// TIA Portal V20 export
FUNCTION_BLOCK "PR_Gantry_2_Soft2.0 1_workflow_0f74f7"   // FB44, LAD
{ S7_Optimized_Access := 'TRUE' }
// stored: MemoryReserve 100, SetENOAutomatically false
   VAR_INPUT
      iAcceptPartPick : Bool;
      iAcceptPartPlace : Bool;
      iAutoRunning : Bool;
      iFaultReset : Bool;
      iFibroSafe : Bool;
      iOTS_Frm_Shuttle : Bool;
      iPartPresent : Bool;
      iPartPresent_Fibro : Bool;
      iPartUngrip : Bool;
      iRTR_Frm_Fibro : Bool;
      iReset_fault : Bool;
      iShuttleAtPickPos : Bool;
      iShuttleSafe : Bool;
      iSstMode : Bool;
      iSstPB : Bool;
      iXAxisAtPartPickPos : Bool;
      iXAxisAtPlacePos : Bool;
      iXAxisSafe : Bool;
      iZAxisDownPlace : Bool;
      iZAxisPickPos : Bool;
      iZAxisSafe : Bool;
      iZAxisUp : Bool;
   END_VAR
   VAR_OUTPUT
      qError : Array[0..8] of Bool;
      qMessage : Array[0..1] of Bool;
      qOTS_To_Fibro : Bool;
      qPartUngripCmd : Bool;
      qRTR_To_Shuttle : Bool;
      qXAxisHomeCmd : Bool;
      qXAxisHomeCmdPlace : Bool;
      qXAxisPickPosCmd : Bool;
      qZAxisDownCmd : Bool;
      qZAxisHomeCmd : Bool;
      qZAxisUpCmd : Bool;
      qZDownCmd : Bool;
   END_VAR
   VAR
      c170_ChkPartPlaced_T1 : Bool;
      c170_ChkPartPlaced_T2 : Bool;
      c180_WtOperatorDecisionPlace_T1 : Bool;
      c180_WtOperatorDecisionPlace_T2 : Bool;
      c40_ChkPartPresent_T1 : Bool;
      c40_ChkPartPresent_T2 : Bool;
      c40_ChkPartPresent_T3 : Bool;
      c90_ChkPartPick_T1 : Bool;
      c90_ChkPartPick_T2 : Bool;
      StateNo : Int;
      s100_WtOperatorDecision : Bool;
      s100_WtOperatorDecision_T1 : Bool;
      s100_WtOperatorDecision_T2 : Bool;
      s10_WtAllAtSafe : Bool;
      s10_WtAllAtSafe_T1 : Bool;
      s110_WtZAxisUp : Bool;
      s110_WtZAxisUp_T1 : Bool;
      s120_ChkFibroSafe : Bool;
      s120_ChkFibroSafe_T1 : Bool;
      s130_WtXAxisPlacePos : Bool;
      s130_WtXAxisPlacePos_T1 : Bool;
      s140_WtRTRFrmFibro : Bool;
      s140_WtRTRFrmFibro_T1 : Bool;
      s150_WtZAxisDownPlace : Bool;
      s150_WtZAxisDownPlace_T1 : Bool;
      s160_WtPartUngrip : Bool;
      s160_WtPartUngrip_T1 : Bool;
      s170_ChkPartPlaced : Bool;
      s170_ChkPartPlaced_T1 : Bool;
      s170_ChkPartPlaced_T2 : Bool;
      s180_WtOperatorDecisionPlace : Bool;
      s180_WtOperatorDecisionPlace_T1 : Bool;
      s180_WtOperatorDecisionPlace_T2 : Bool;
      s1_ResetRelease : Bool;
      s1_ResetRelease_T1 : Bool;
      s20_WtZAxisSafe : Bool;
      s20_WtZAxisSafe_T1 : Bool;
      s30_WtXAxisAtSafe : Bool;
      s30_WtXAxisAtSafe_T1 : Bool;
      s40_ChkPartPresent : Bool;
      s40_ChkPartPresent_T1 : Bool;
      s40_ChkPartPresent_T2 : Bool;
      s40_ChkPartPresent_T3 : Bool;
      s45_WtOperatorAck : Bool;
      s45_WtOperatorAck_T1 : Bool;
      s50_WtShuttleAtSafe : Bool;
      s50_WtShuttleAtSafe_T1 : Bool;
      s60_WtXAxisPickPos : Bool;
      s60_WtXAxisPickPos_T1 : Bool;
      s70_WtOTSFrmShuttle : Bool;
      s70_WtOTSFrmShuttle_T1 : Bool;
      s80_WtZAxisPickPos : Bool;
      s80_WtZAxisPickPos_T1 : Bool;
      s90_ChkPartPick : Bool;
      s90_ChkPartPick_T1 : Bool;
      s90_ChkPartPick_T2 : Bool;
      sAbnormalStatus : Bool;
      sPartPresentInGrip : Bool;
      sSst : Bool;
      sSstPulse : Bool;
      sSstRise : Bool;
      sStWtResetRel : Bool;
      sStWtResetRel_T1 : Bool;
   END_VAR
   VAR_TEMP
      tOne : Bool;
   END_VAR
   VAR_TEMP   // added for the SCL form of the ladder/FBD networks
      _w1 : Bool;
      _w2 : Bool;
   END_VAR
BEGIN

REGION Network 1
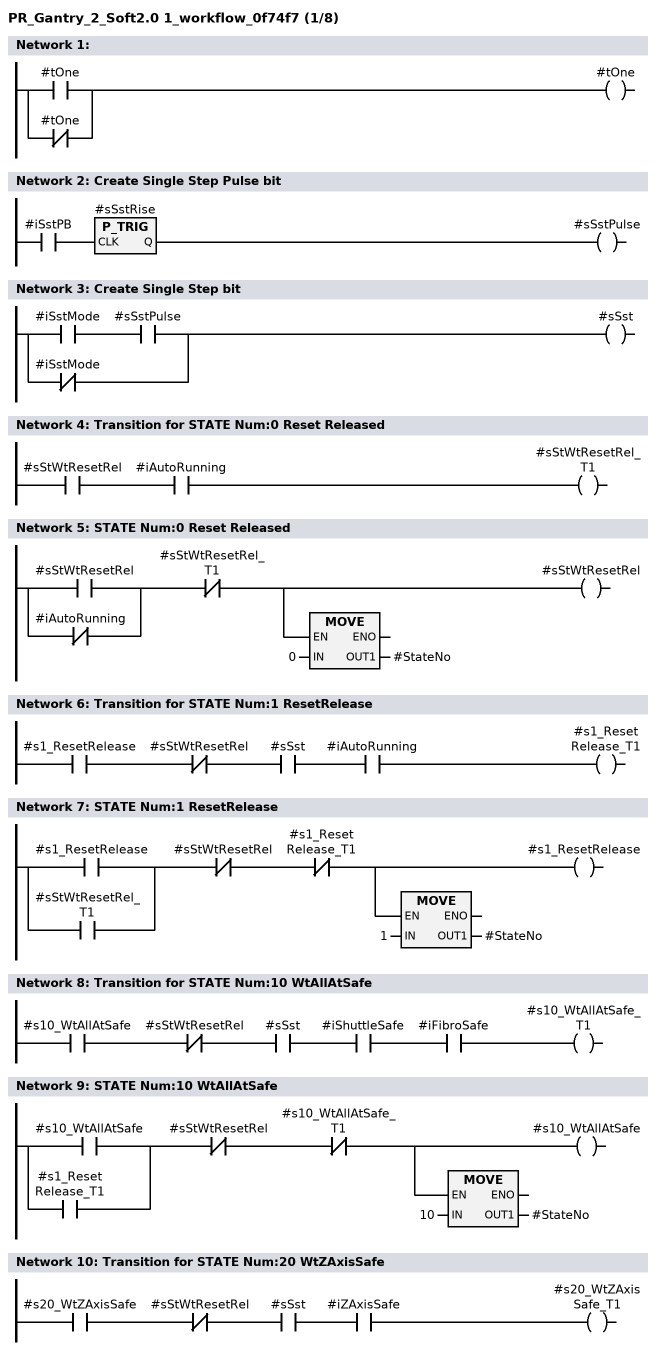
   RUNG wire#powerrail
      Contact( #tOne )
      wire#w1
      Coil( #tOne )
   END_RUNG
   RUNG wire#powerrail
      I_Contact( #tOne )
   END_RUNG wire#w1
   // the same network as SCL:
   #tOne := #tOne OR NOT #tOne;
END_REGION

REGION Network 2: Create Single Step Pulse bit
   RUNG wire#powerrail
      Contact( #iSstPB )
      P_Trig( #sSstRise )
      Coil( #sSstPulse )
   END_RUNG
   // the same network as SCL:
   #_w1 := #iSstPB AND NOT #sSstRise;   // rising edge
   #sSstRise := #iSstPB;
   #sSstPulse := #_w1;
END_REGION

REGION Network 3: Create Single Step bit
   RUNG wire#powerrail
      Contact( #iSstMode )
      Contact( #sSstPulse )
      wire#w1
      Coil( #sSst )
   END_RUNG
   RUNG wire#powerrail
      I_Contact( #iSstMode )
   END_RUNG wire#w1
   // the same network as SCL:
   #sSst := (#iSstMode AND #sSstPulse) OR NOT #iSstMode;
END_REGION

REGION Network 4: Transition for STATE Num:0 Reset Released
   RUNG wire#powerrail
      Contact( #sStWtResetRel )
      Contact( #iAutoRunning )
      Coil( #sStWtResetRel_T1 )
   END_RUNG
   // the same network as SCL:
   #sStWtResetRel_T1 := #sStWtResetRel AND #iAutoRunning;
END_REGION

REGION Network 5: STATE Num:0 Reset Released
   RUNG wire#powerrail
      Contact( #sStWtResetRel )
      wire#w1
      I_Contact( #sStWtResetRel_T1 )
      wire#w2
      Coil( #sStWtResetRel )
   END_RUNG
   RUNG wire#powerrail
      I_Contact( #iAutoRunning )
   END_RUNG wire#w1
   RUNG wire#w2
      { S7_GenerateENO := "TRUE" } Move(in := 0, out1 => #StateNo)
   END_RUNG
   // the same network as SCL:
   #sStWtResetRel := (#sStWtResetRel OR NOT #iAutoRunning) AND NOT #sStWtResetRel_T1;
   IF #sStWtResetRel THEN #StateNo := 0; END_IF;
END_REGION

REGION Network 6: Transition for STATE Num:1 ResetRelease
   RUNG wire#powerrail
      Contact( #s1_ResetRelease )
      I_Contact( #sStWtResetRel )
      Contact( #sSst )
      Contact( #iAutoRunning )
      Coil( #s1_ResetRelease_T1 )
   END_RUNG
   // the same network as SCL:
   #s1_ResetRelease_T1 := #s1_ResetRelease AND NOT #sStWtResetRel AND #sSst AND #iAutoRunning;
END_REGION

REGION Network 7: STATE Num:1 ResetRelease
   RUNG wire#powerrail
      Contact( #s1_ResetRelease )
      wire#w1
      I_Contact( #sStWtResetRel )
      I_Contact( #s1_ResetRelease_T1 )
      wire#w2
      Coil( #s1_ResetRelease )
   END_RUNG
   RUNG wire#powerrail
      Contact( #sStWtResetRel_T1 )
   END_RUNG wire#w1
   RUNG wire#w2
      { S7_GenerateENO := "TRUE" } Move(in := 1, out1 => #StateNo)
   END_RUNG
   // the same network as SCL:
   #s1_ResetRelease := (#s1_ResetRelease OR #sStWtResetRel_T1) AND NOT #sStWtResetRel AND NOT #s1_ResetRelease_T1;
   IF #s1_ResetRelease THEN #StateNo := 1; END_IF;
END_REGION

REGION Network 8: Transition for STATE Num:10 WtAllAtSafe
   RUNG wire#powerrail
      Contact( #s10_WtAllAtSafe )
      I_Contact( #sStWtResetRel )
      Contact( #sSst )
      Contact( #iShuttleSafe )
      Contact( #iFibroSafe )
      Coil( #s10_WtAllAtSafe_T1 )
   END_RUNG
   // the same network as SCL:
   #s10_WtAllAtSafe_T1 := #s10_WtAllAtSafe AND NOT #sStWtResetRel AND #sSst AND #iShuttleSafe AND #iFibroSafe;
END_REGION

REGION Network 9: STATE Num:10 WtAllAtSafe
   RUNG wire#powerrail
      Contact( #s10_WtAllAtSafe )
      wire#w1
      I_Contact( #sStWtResetRel )
      I_Contact( #s10_WtAllAtSafe_T1 )
      wire#w2
      Coil( #s10_WtAllAtSafe )
   END_RUNG
   RUNG wire#powerrail
      Contact( #s1_ResetRelease_T1 )
   END_RUNG wire#w1
   RUNG wire#w2
      { S7_GenerateENO := "TRUE" } Move(in := 10, out1 => #StateNo)
   END_RUNG
   // the same network as SCL:
   #s10_WtAllAtSafe := (#s10_WtAllAtSafe OR #s1_ResetRelease_T1) AND NOT #sStWtResetRel AND NOT #s10_WtAllAtSafe_T1;
   IF #s10_WtAllAtSafe THEN #StateNo := 10; END_IF;
END_REGION

REGION Network 10: Transition for STATE Num:20 WtZAxisSafe
   RUNG wire#powerrail
      Contact( #s20_WtZAxisSafe )
      I_Contact( #sStWtResetRel )
      Contact( #sSst )
      Contact( #iZAxisSafe )
      Coil( #s20_WtZAxisSafe_T1 )
   END_RUNG
   // the same network as SCL:
   #s20_WtZAxisSafe_T1 := #s20_WtZAxisSafe AND NOT #sStWtResetRel AND #sSst AND #iZAxisSafe;
END_REGION

REGION Network 11: STATE Num:20 WtZAxisSafe
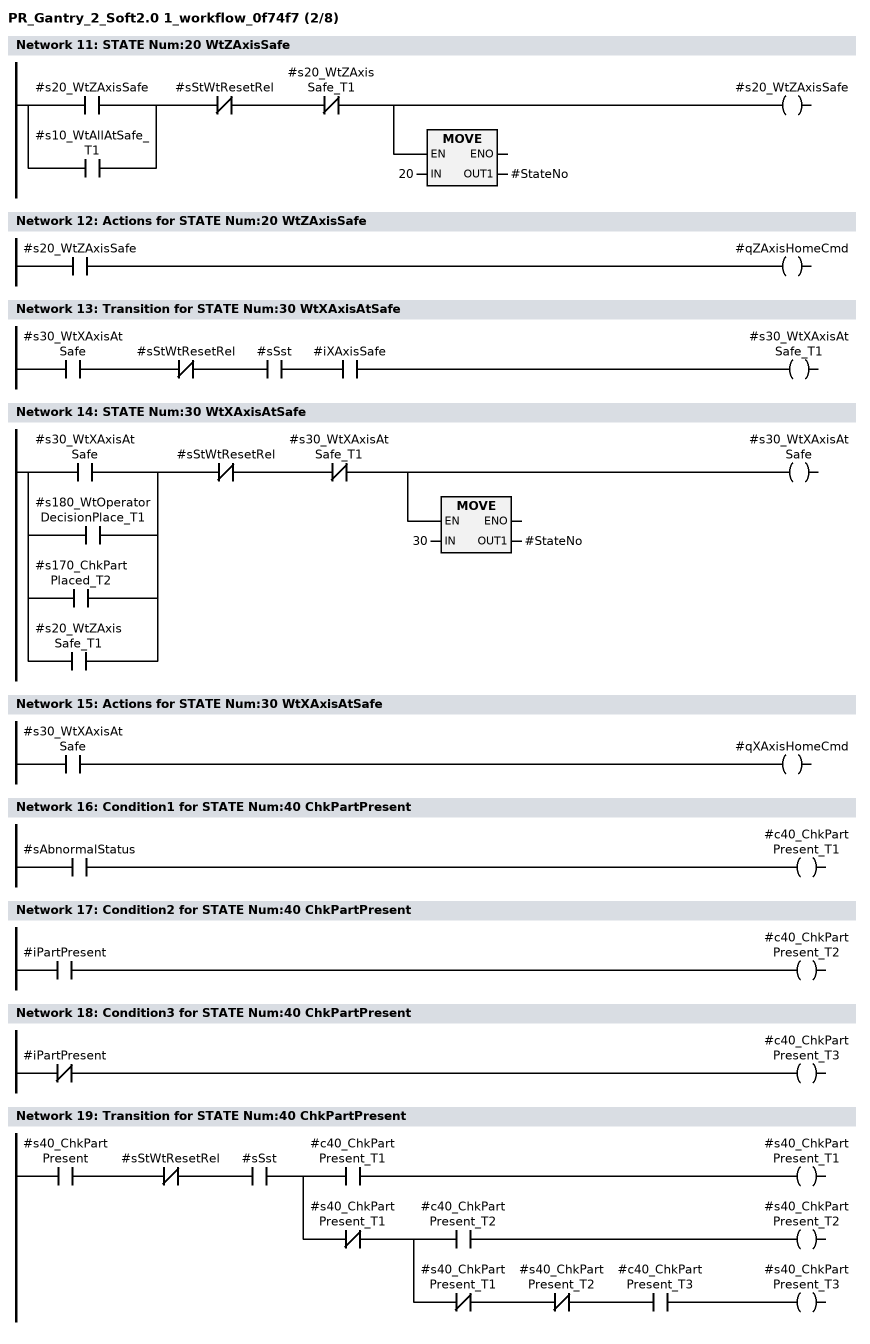
   RUNG wire#powerrail
      Contact( #s20_WtZAxisSafe )
      wire#w1
      I_Contact( #sStWtResetRel )
      I_Contact( #s20_WtZAxisSafe_T1 )
      wire#w2
      Coil( #s20_WtZAxisSafe )
   END_RUNG
   RUNG wire#powerrail
      Contact( #s10_WtAllAtSafe_T1 )
   END_RUNG wire#w1
   RUNG wire#w2
      { S7_GenerateENO := "TRUE" } Move(in := 20, out1 => #StateNo)
   END_RUNG
   // the same network as SCL:
   #s20_WtZAxisSafe := (#s20_WtZAxisSafe OR #s10_WtAllAtSafe_T1) AND NOT #sStWtResetRel AND NOT #s20_WtZAxisSafe_T1;
   IF #s20_WtZAxisSafe THEN #StateNo := 20; END_IF;
END_REGION

REGION Network 12: Actions for STATE Num:20 WtZAxisSafe
   RUNG wire#powerrail
      Contact( #s20_WtZAxisSafe )
      Coil( #qZAxisHomeCmd )
   END_RUNG
   // the same network as SCL:
   #qZAxisHomeCmd := #s20_WtZAxisSafe;
END_REGION

REGION Network 13: Transition for STATE Num:30 WtXAxisAtSafe
   RUNG wire#powerrail
      Contact( #s30_WtXAxisAtSafe )
      I_Contact( #sStWtResetRel )
      Contact( #sSst )
      Contact( #iXAxisSafe )
      Coil( #s30_WtXAxisAtSafe_T1 )
   END_RUNG
   // the same network as SCL:
   #s30_WtXAxisAtSafe_T1 := #s30_WtXAxisAtSafe AND NOT #sStWtResetRel AND #sSst AND #iXAxisSafe;
END_REGION

REGION Network 14: STATE Num:30 WtXAxisAtSafe
   RUNG wire#powerrail
      Contact( #s30_WtXAxisAtSafe )
      wire#w1
      I_Contact( #sStWtResetRel )
      I_Contact( #s30_WtXAxisAtSafe_T1 )
      wire#w2
      Coil( #s30_WtXAxisAtSafe )
   END_RUNG
   RUNG wire#powerrail
      Contact( #s180_WtOperatorDecisionPlace_T1 )
   END_RUNG wire#w1
   RUNG wire#powerrail
      Contact( #s170_ChkPartPlaced_T2 )
   END_RUNG wire#w1
   RUNG wire#powerrail
      Contact( #s20_WtZAxisSafe_T1 )
   END_RUNG wire#w1
   RUNG wire#w2
      { S7_GenerateENO := "TRUE" } Move(in := 30, out1 => #StateNo)
   END_RUNG
   // the same network as SCL:
   #s30_WtXAxisAtSafe := (#s30_WtXAxisAtSafe OR #s180_WtOperatorDecisionPlace_T1 OR #s170_ChkPartPlaced_T2 OR #s20_WtZAxisSafe_T1) AND NOT #sStWtResetRel AND NOT #s30_WtXAxisAtSafe_T1;
   IF #s30_WtXAxisAtSafe THEN #StateNo := 30; END_IF;
END_REGION

REGION Network 15: Actions for STATE Num:30 WtXAxisAtSafe
   RUNG wire#powerrail
      Contact( #s30_WtXAxisAtSafe )
      Coil( #qXAxisHomeCmd )
   END_RUNG
   // the same network as SCL:
   #qXAxisHomeCmd := #s30_WtXAxisAtSafe;
END_REGION

REGION Network 16: Condition1 for STATE Num:40 ChkPartPresent
   RUNG wire#powerrail
      Contact( #sAbnormalStatus )
      Coil( #c40_ChkPartPresent_T1 )
   END_RUNG
   // the same network as SCL:
   #c40_ChkPartPresent_T1 := #sAbnormalStatus;
END_REGION

REGION Network 17: Condition2 for STATE Num:40 ChkPartPresent
   RUNG wire#powerrail
      Contact( #iPartPresent )
      Coil( #c40_ChkPartPresent_T2 )
   END_RUNG
   // the same network as SCL:
   #c40_ChkPartPresent_T2 := #iPartPresent;
END_REGION

REGION Network 18: Condition3 for STATE Num:40 ChkPartPresent
   RUNG wire#powerrail
      I_Contact( #iPartPresent )
      Coil( #c40_ChkPartPresent_T3 )
   END_RUNG
   // the same network as SCL:
   #c40_ChkPartPresent_T3 := NOT #iPartPresent;
END_REGION

REGION Network 19: Transition for STATE Num:40 ChkPartPresent
   RUNG wire#powerrail
      Contact( #s40_ChkPartPresent )
      I_Contact( #sStWtResetRel )
      Contact( #sSst )
      wire#w1
      Contact( #c40_ChkPartPresent_T1 )
      Coil( #s40_ChkPartPresent_T1 )
   END_RUNG
   RUNG wire#w1
      I_Contact( #s40_ChkPartPresent_T1 )
      wire#w2
      Contact( #c40_ChkPartPresent_T2 )
      Coil( #s40_ChkPartPresent_T2 )
   END_RUNG
   RUNG wire#w2
      I_Contact( #s40_ChkPartPresent_T1 )
      I_Contact( #s40_ChkPartPresent_T2 )
      Contact( #c40_ChkPartPresent_T3 )
      Coil( #s40_ChkPartPresent_T3 )
   END_RUNG
   // the same network as SCL:
   #_w1 := #s40_ChkPartPresent AND NOT #sStWtResetRel AND #sSst;
   #s40_ChkPartPresent_T1 := #_w1 AND #c40_ChkPartPresent_T1;
   #_w2 := #_w1 AND NOT #s40_ChkPartPresent_T1;
   #s40_ChkPartPresent_T2 := #_w2 AND #c40_ChkPartPresent_T2;
   #s40_ChkPartPresent_T3 := #_w2 AND NOT #s40_ChkPartPresent_T1 AND NOT #s40_ChkPartPresent_T2 AND #c40_ChkPartPresent_T3;
END_REGION

REGION Network 20: STATE Num:40 ChkPartPresent
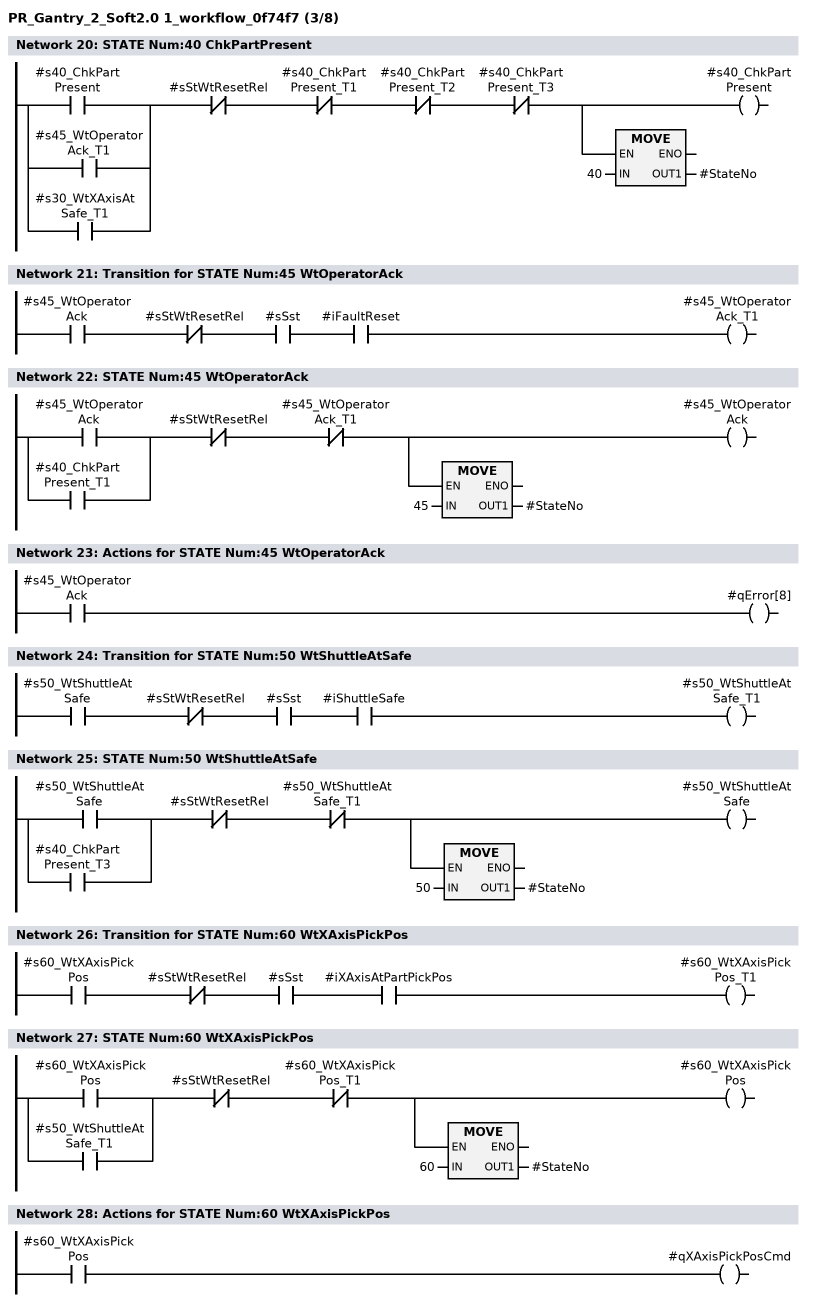
   RUNG wire#powerrail
      Contact( #s40_ChkPartPresent )
      wire#w1
      I_Contact( #sStWtResetRel )
      I_Contact( #s40_ChkPartPresent_T1 )
      I_Contact( #s40_ChkPartPresent_T2 )
      I_Contact( #s40_ChkPartPresent_T3 )
      wire#w2
      Coil( #s40_ChkPartPresent )
   END_RUNG
   RUNG wire#powerrail
      Contact( #s45_WtOperatorAck_T1 )
   END_RUNG wire#w1
   RUNG wire#powerrail
      Contact( #s30_WtXAxisAtSafe_T1 )
   END_RUNG wire#w1
   RUNG wire#w2
      { S7_GenerateENO := "TRUE" } Move(in := 40, out1 => #StateNo)
   END_RUNG
   // the same network as SCL:
   #s40_ChkPartPresent := (#s40_ChkPartPresent OR #s45_WtOperatorAck_T1 OR #s30_WtXAxisAtSafe_T1) AND NOT #sStWtResetRel AND NOT #s40_ChkPartPresent_T1 AND NOT #s40_ChkPartPresent_T2 AND NOT #s40_ChkPartPresent_T3;
   IF #s40_ChkPartPresent THEN #StateNo := 40; END_IF;
END_REGION

REGION Network 21: Transition for STATE Num:45 WtOperatorAck
   RUNG wire#powerrail
      Contact( #s45_WtOperatorAck )
      I_Contact( #sStWtResetRel )
      Contact( #sSst )
      Contact( #iFaultReset )
      Coil( #s45_WtOperatorAck_T1 )
   END_RUNG
   // the same network as SCL:
   #s45_WtOperatorAck_T1 := #s45_WtOperatorAck AND NOT #sStWtResetRel AND #sSst AND #iFaultReset;
END_REGION

REGION Network 22: STATE Num:45 WtOperatorAck
   RUNG wire#powerrail
      Contact( #s45_WtOperatorAck )
      wire#w1
      I_Contact( #sStWtResetRel )
      I_Contact( #s45_WtOperatorAck_T1 )
      wire#w2
      Coil( #s45_WtOperatorAck )
   END_RUNG
   RUNG wire#powerrail
      Contact( #s40_ChkPartPresent_T1 )
   END_RUNG wire#w1
   RUNG wire#w2
      { S7_GenerateENO := "TRUE" } Move(in := 45, out1 => #StateNo)
   END_RUNG
   // the same network as SCL:
   #s45_WtOperatorAck := (#s45_WtOperatorAck OR #s40_ChkPartPresent_T1) AND NOT #sStWtResetRel AND NOT #s45_WtOperatorAck_T1;
   IF #s45_WtOperatorAck THEN #StateNo := 45; END_IF;
END_REGION

REGION Network 23: Actions for STATE Num:45 WtOperatorAck
   RUNG wire#powerrail
      Contact( #s45_WtOperatorAck )
      Coil( #qError[8] )
   END_RUNG
   // the same network as SCL:
   #qError[8] := #s45_WtOperatorAck;
END_REGION

REGION Network 24: Transition for STATE Num:50 WtShuttleAtSafe
   RUNG wire#powerrail
      Contact( #s50_WtShuttleAtSafe )
      I_Contact( #sStWtResetRel )
      Contact( #sSst )
      Contact( #iShuttleSafe )
      Coil( #s50_WtShuttleAtSafe_T1 )
   END_RUNG
   // the same network as SCL:
   #s50_WtShuttleAtSafe_T1 := #s50_WtShuttleAtSafe AND NOT #sStWtResetRel AND #sSst AND #iShuttleSafe;
END_REGION

REGION Network 25: STATE Num:50 WtShuttleAtSafe
   RUNG wire#powerrail
      Contact( #s50_WtShuttleAtSafe )
      wire#w1
      I_Contact( #sStWtResetRel )
      I_Contact( #s50_WtShuttleAtSafe_T1 )
      wire#w2
      Coil( #s50_WtShuttleAtSafe )
   END_RUNG
   RUNG wire#powerrail
      Contact( #s40_ChkPartPresent_T3 )
   END_RUNG wire#w1
   RUNG wire#w2
      { S7_GenerateENO := "TRUE" } Move(in := 50, out1 => #StateNo)
   END_RUNG
   // the same network as SCL:
   #s50_WtShuttleAtSafe := (#s50_WtShuttleAtSafe OR #s40_ChkPartPresent_T3) AND NOT #sStWtResetRel AND NOT #s50_WtShuttleAtSafe_T1;
   IF #s50_WtShuttleAtSafe THEN #StateNo := 50; END_IF;
END_REGION

REGION Network 26: Transition for STATE Num:60 WtXAxisPickPos
   RUNG wire#powerrail
      Contact( #s60_WtXAxisPickPos )
      I_Contact( #sStWtResetRel )
      Contact( #sSst )
      Contact( #iXAxisAtPartPickPos )
      Coil( #s60_WtXAxisPickPos_T1 )
   END_RUNG
   // the same network as SCL:
   #s60_WtXAxisPickPos_T1 := #s60_WtXAxisPickPos AND NOT #sStWtResetRel AND #sSst AND #iXAxisAtPartPickPos;
END_REGION

REGION Network 27: STATE Num:60 WtXAxisPickPos
   RUNG wire#powerrail
      Contact( #s60_WtXAxisPickPos )
      wire#w1
      I_Contact( #sStWtResetRel )
      I_Contact( #s60_WtXAxisPickPos_T1 )
      wire#w2
      Coil( #s60_WtXAxisPickPos )
   END_RUNG
   RUNG wire#powerrail
      Contact( #s50_WtShuttleAtSafe_T1 )
   END_RUNG wire#w1
   RUNG wire#w2
      { S7_GenerateENO := "TRUE" } Move(in := 60, out1 => #StateNo)
   END_RUNG
   // the same network as SCL:
   #s60_WtXAxisPickPos := (#s60_WtXAxisPickPos OR #s50_WtShuttleAtSafe_T1) AND NOT #sStWtResetRel AND NOT #s60_WtXAxisPickPos_T1;
   IF #s60_WtXAxisPickPos THEN #StateNo := 60; END_IF;
END_REGION

REGION Network 28: Actions for STATE Num:60 WtXAxisPickPos
   RUNG wire#powerrail
      Contact( #s60_WtXAxisPickPos )
      Coil( #qXAxisPickPosCmd )
   END_RUNG
   // the same network as SCL:
   #qXAxisPickPosCmd := #s60_WtXAxisPickPos;
END_REGION

REGION Network 29: Transition for STATE Num:70 WtOTSFrmShuttle
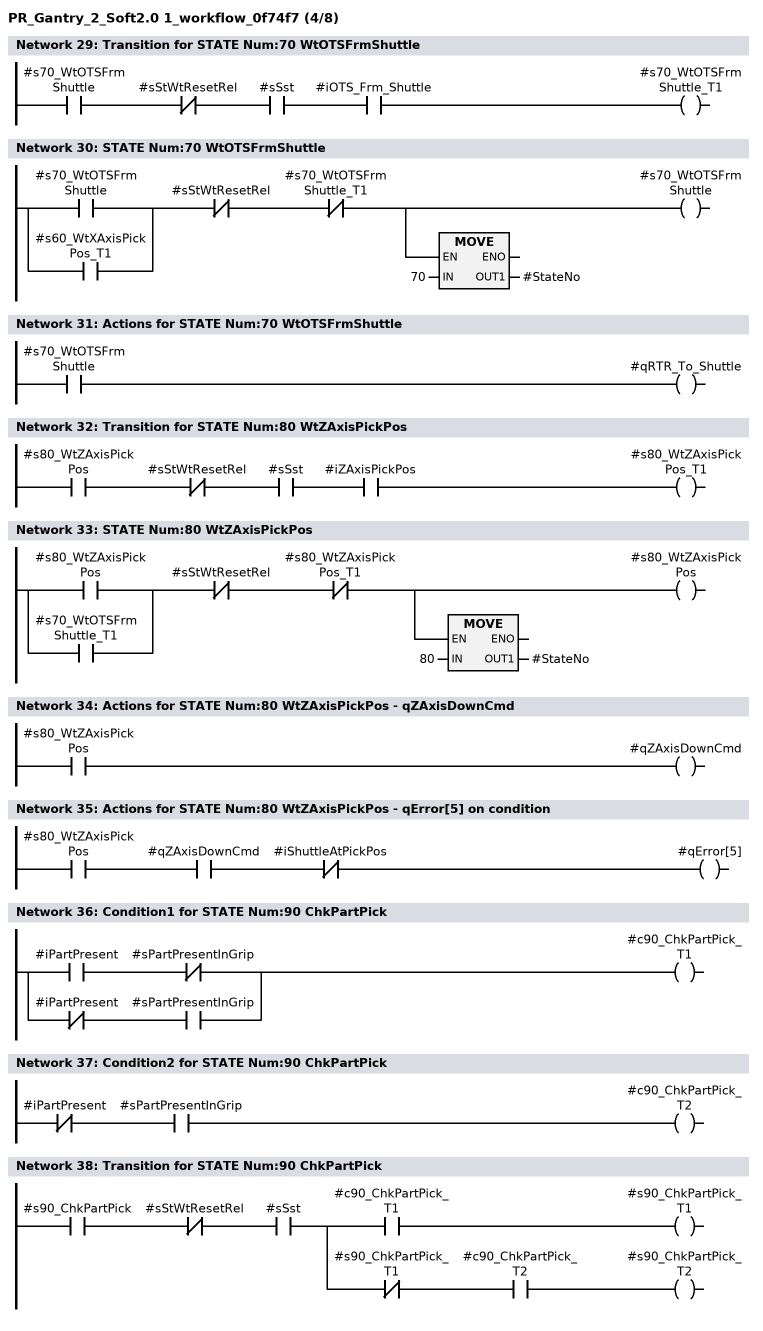
   RUNG wire#powerrail
      Contact( #s70_WtOTSFrmShuttle )
      I_Contact( #sStWtResetRel )
      Contact( #sSst )
      Contact( #iOTS_Frm_Shuttle )
      Coil( #s70_WtOTSFrmShuttle_T1 )
   END_RUNG
   // the same network as SCL:
   #s70_WtOTSFrmShuttle_T1 := #s70_WtOTSFrmShuttle AND NOT #sStWtResetRel AND #sSst AND #iOTS_Frm_Shuttle;
END_REGION

REGION Network 30: STATE Num:70 WtOTSFrmShuttle
   RUNG wire#powerrail
      Contact( #s70_WtOTSFrmShuttle )
      wire#w1
      I_Contact( #sStWtResetRel )
      I_Contact( #s70_WtOTSFrmShuttle_T1 )
      wire#w2
      Coil( #s70_WtOTSFrmShuttle )
   END_RUNG
   RUNG wire#powerrail
      Contact( #s60_WtXAxisPickPos_T1 )
   END_RUNG wire#w1
   RUNG wire#w2
      { S7_GenerateENO := "TRUE" } Move(in := 70, out1 => #StateNo)
   END_RUNG
   // the same network as SCL:
   #s70_WtOTSFrmShuttle := (#s70_WtOTSFrmShuttle OR #s60_WtXAxisPickPos_T1) AND NOT #sStWtResetRel AND NOT #s70_WtOTSFrmShuttle_T1;
   IF #s70_WtOTSFrmShuttle THEN #StateNo := 70; END_IF;
END_REGION

REGION Network 31: Actions for STATE Num:70 WtOTSFrmShuttle
   RUNG wire#powerrail
      Contact( #s70_WtOTSFrmShuttle )
      Coil( #qRTR_To_Shuttle )
   END_RUNG
   // the same network as SCL:
   #qRTR_To_Shuttle := #s70_WtOTSFrmShuttle;
END_REGION

REGION Network 32: Transition for STATE Num:80 WtZAxisPickPos
   RUNG wire#powerrail
      Contact( #s80_WtZAxisPickPos )
      I_Contact( #sStWtResetRel )
      Contact( #sSst )
      Contact( #iZAxisPickPos )
      Coil( #s80_WtZAxisPickPos_T1 )
   END_RUNG
   // the same network as SCL:
   #s80_WtZAxisPickPos_T1 := #s80_WtZAxisPickPos AND NOT #sStWtResetRel AND #sSst AND #iZAxisPickPos;
END_REGION

REGION Network 33: STATE Num:80 WtZAxisPickPos
   RUNG wire#powerrail
      Contact( #s80_WtZAxisPickPos )
      wire#w1
      I_Contact( #sStWtResetRel )
      I_Contact( #s80_WtZAxisPickPos_T1 )
      wire#w2
      Coil( #s80_WtZAxisPickPos )
   END_RUNG
   RUNG wire#powerrail
      Contact( #s70_WtOTSFrmShuttle_T1 )
   END_RUNG wire#w1
   RUNG wire#w2
      { S7_GenerateENO := "TRUE" } Move(in := 80, out1 => #StateNo)
   END_RUNG
   // the same network as SCL:
   #s80_WtZAxisPickPos := (#s80_WtZAxisPickPos OR #s70_WtOTSFrmShuttle_T1) AND NOT #sStWtResetRel AND NOT #s80_WtZAxisPickPos_T1;
   IF #s80_WtZAxisPickPos THEN #StateNo := 80; END_IF;
END_REGION

REGION Network 34: Actions for STATE Num:80 WtZAxisPickPos - qZAxisDownCmd
   RUNG wire#powerrail
      Contact( #s80_WtZAxisPickPos )
      Coil( #qZAxisDownCmd )
   END_RUNG
   // the same network as SCL:
   #qZAxisDownCmd := #s80_WtZAxisPickPos;
END_REGION

REGION Network 35: Actions for STATE Num:80 WtZAxisPickPos - qError[5] on condition
   RUNG wire#powerrail
      Contact( #s80_WtZAxisPickPos )
      Contact( #qZAxisDownCmd )
      I_Contact( #iShuttleAtPickPos )
      Coil( #qError[5] )
   END_RUNG
   // the same network as SCL:
   #qError[5] := #s80_WtZAxisPickPos AND #qZAxisDownCmd AND NOT #iShuttleAtPickPos;
END_REGION

REGION Network 36: Condition1 for STATE Num:90 ChkPartPick
   RUNG wire#powerrail
      Contact( #iPartPresent )
      I_Contact( #sPartPresentInGrip )
      wire#w1
      Coil( #c90_ChkPartPick_T1 )
   END_RUNG
   RUNG wire#powerrail
      I_Contact( #iPartPresent )
      Contact( #sPartPresentInGrip )
   END_RUNG wire#w1
   // the same network as SCL:
   #c90_ChkPartPick_T1 := (#iPartPresent AND NOT #sPartPresentInGrip) OR (NOT #iPartPresent AND #sPartPresentInGrip);
END_REGION

REGION Network 37: Condition2 for STATE Num:90 ChkPartPick
   RUNG wire#powerrail
      I_Contact( #iPartPresent )
      Contact( #sPartPresentInGrip )
      Coil( #c90_ChkPartPick_T2 )
   END_RUNG
   // the same network as SCL:
   #c90_ChkPartPick_T2 := NOT #iPartPresent AND #sPartPresentInGrip;
END_REGION

REGION Network 38: Transition for STATE Num:90 ChkPartPick
   RUNG wire#powerrail
      Contact( #s90_ChkPartPick )
      I_Contact( #sStWtResetRel )
      Contact( #sSst )
      wire#w1
      Contact( #c90_ChkPartPick_T1 )
      Coil( #s90_ChkPartPick_T1 )
   END_RUNG
   RUNG wire#w1
      I_Contact( #s90_ChkPartPick_T1 )
      Contact( #c90_ChkPartPick_T2 )
      Coil( #s90_ChkPartPick_T2 )
   END_RUNG
   // the same network as SCL:
   #_w1 := #s90_ChkPartPick AND NOT #sStWtResetRel AND #sSst;
   #s90_ChkPartPick_T1 := #_w1 AND #c90_ChkPartPick_T1;
   #s90_ChkPartPick_T2 := #_w1 AND NOT #s90_ChkPartPick_T1 AND #c90_ChkPartPick_T2;
END_REGION

REGION Network 39: STATE Num:90 ChkPartPick
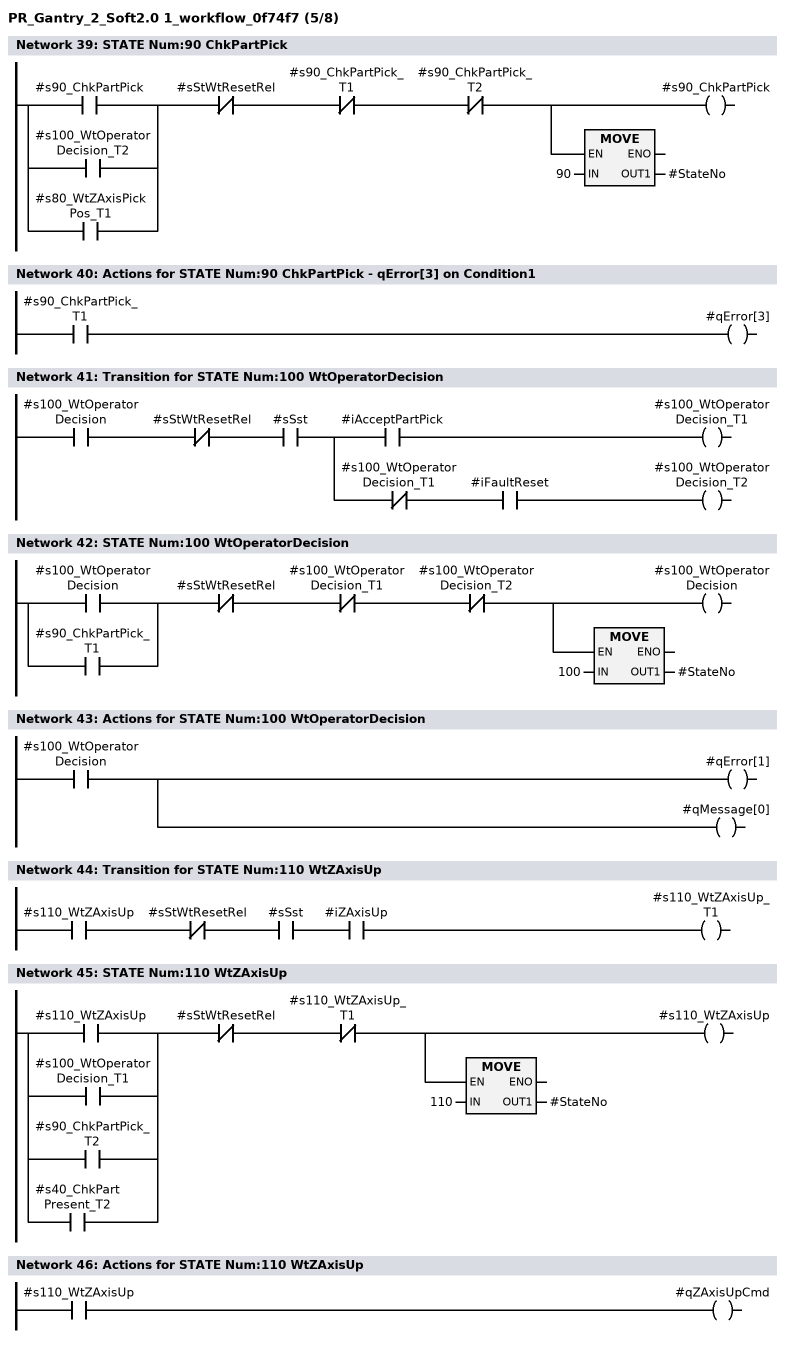
   RUNG wire#powerrail
      Contact( #s90_ChkPartPick )
      wire#w1
      I_Contact( #sStWtResetRel )
      I_Contact( #s90_ChkPartPick_T1 )
      I_Contact( #s90_ChkPartPick_T2 )
      wire#w2
      Coil( #s90_ChkPartPick )
   END_RUNG
   RUNG wire#powerrail
      Contact( #s100_WtOperatorDecision_T2 )
   END_RUNG wire#w1
   RUNG wire#powerrail
      Contact( #s80_WtZAxisPickPos_T1 )
   END_RUNG wire#w1
   RUNG wire#w2
      { S7_GenerateENO := "TRUE" } Move(in := 90, out1 => #StateNo)
   END_RUNG
   // the same network as SCL:
   #s90_ChkPartPick := (#s90_ChkPartPick OR #s100_WtOperatorDecision_T2 OR #s80_WtZAxisPickPos_T1) AND NOT #sStWtResetRel AND NOT #s90_ChkPartPick_T1 AND NOT #s90_ChkPartPick_T2;
   IF #s90_ChkPartPick THEN #StateNo := 90; END_IF;
END_REGION

REGION Network 40: Actions for STATE Num:90 ChkPartPick - qError[3] on Condition1
   RUNG wire#powerrail
      Contact( #s90_ChkPartPick_T1 )
      Coil( #qError[3] )
   END_RUNG
   // the same network as SCL:
   #qError[3] := #s90_ChkPartPick_T1;
END_REGION

REGION Network 41: Transition for STATE Num:100 WtOperatorDecision
   RUNG wire#powerrail
      Contact( #s100_WtOperatorDecision )
      I_Contact( #sStWtResetRel )
      Contact( #sSst )
      wire#w1
      Contact( #iAcceptPartPick )
      Coil( #s100_WtOperatorDecision_T1 )
   END_RUNG
   RUNG wire#w1
      I_Contact( #s100_WtOperatorDecision_T1 )
      Contact( #iFaultReset )
      Coil( #s100_WtOperatorDecision_T2 )
   END_RUNG
   // the same network as SCL:
   #_w1 := #s100_WtOperatorDecision AND NOT #sStWtResetRel AND #sSst;
   #s100_WtOperatorDecision_T1 := #_w1 AND #iAcceptPartPick;
   #s100_WtOperatorDecision_T2 := #_w1 AND NOT #s100_WtOperatorDecision_T1 AND #iFaultReset;
END_REGION

REGION Network 42: STATE Num:100 WtOperatorDecision
   RUNG wire#powerrail
      Contact( #s100_WtOperatorDecision )
      wire#w1
      I_Contact( #sStWtResetRel )
      I_Contact( #s100_WtOperatorDecision_T1 )
      I_Contact( #s100_WtOperatorDecision_T2 )
      wire#w2
      Coil( #s100_WtOperatorDecision )
   END_RUNG
   RUNG wire#powerrail
      Contact( #s90_ChkPartPick_T1 )
   END_RUNG wire#w1
   RUNG wire#w2
      { S7_GenerateENO := "TRUE" } Move(in := 100, out1 => #StateNo)
   END_RUNG
   // the same network as SCL:
   #s100_WtOperatorDecision := (#s100_WtOperatorDecision OR #s90_ChkPartPick_T1) AND NOT #sStWtResetRel AND NOT #s100_WtOperatorDecision_T1 AND NOT #s100_WtOperatorDecision_T2;
   IF #s100_WtOperatorDecision THEN #StateNo := 100; END_IF;
END_REGION

REGION Network 43: Actions for STATE Num:100 WtOperatorDecision
   RUNG wire#powerrail
      Contact( #s100_WtOperatorDecision )
      wire#w1
      Coil( #qError[1] )
   END_RUNG
   RUNG wire#w1
      Coil( #qMessage[0] )
   END_RUNG
   // the same network as SCL:
   #qError[1] := #s100_WtOperatorDecision;
   #qMessage[0] := #s100_WtOperatorDecision;
END_REGION

REGION Network 44: Transition for STATE Num:110 WtZAxisUp
   RUNG wire#powerrail
      Contact( #s110_WtZAxisUp )
      I_Contact( #sStWtResetRel )
      Contact( #sSst )
      Contact( #iZAxisUp )
      Coil( #s110_WtZAxisUp_T1 )
   END_RUNG
   // the same network as SCL:
   #s110_WtZAxisUp_T1 := #s110_WtZAxisUp AND NOT #sStWtResetRel AND #sSst AND #iZAxisUp;
END_REGION

REGION Network 45: STATE Num:110 WtZAxisUp
   RUNG wire#powerrail
      Contact( #s110_WtZAxisUp )
      wire#w1
      I_Contact( #sStWtResetRel )
      I_Contact( #s110_WtZAxisUp_T1 )
      wire#w2
      Coil( #s110_WtZAxisUp )
   END_RUNG
   RUNG wire#powerrail
      Contact( #s100_WtOperatorDecision_T1 )
   END_RUNG wire#w1
   RUNG wire#powerrail
      Contact( #s90_ChkPartPick_T2 )
   END_RUNG wire#w1
   RUNG wire#powerrail
      Contact( #s40_ChkPartPresent_T2 )
   END_RUNG wire#w1
   RUNG wire#w2
      { S7_GenerateENO := "TRUE" } Move(in := 110, out1 => #StateNo)
   END_RUNG
   // the same network as SCL:
   #s110_WtZAxisUp := (#s110_WtZAxisUp OR #s100_WtOperatorDecision_T1 OR #s90_ChkPartPick_T2 OR #s40_ChkPartPresent_T2) AND NOT #sStWtResetRel AND NOT #s110_WtZAxisUp_T1;
   IF #s110_WtZAxisUp THEN #StateNo := 110; END_IF;
END_REGION

REGION Network 46: Actions for STATE Num:110 WtZAxisUp
   RUNG wire#powerrail
      Contact( #s110_WtZAxisUp )
      Coil( #qZAxisUpCmd )
   END_RUNG
   // the same network as SCL:
   #qZAxisUpCmd := #s110_WtZAxisUp;
END_REGION

REGION Network 47: Transition for STATE Num:120 ChkFibroSafe
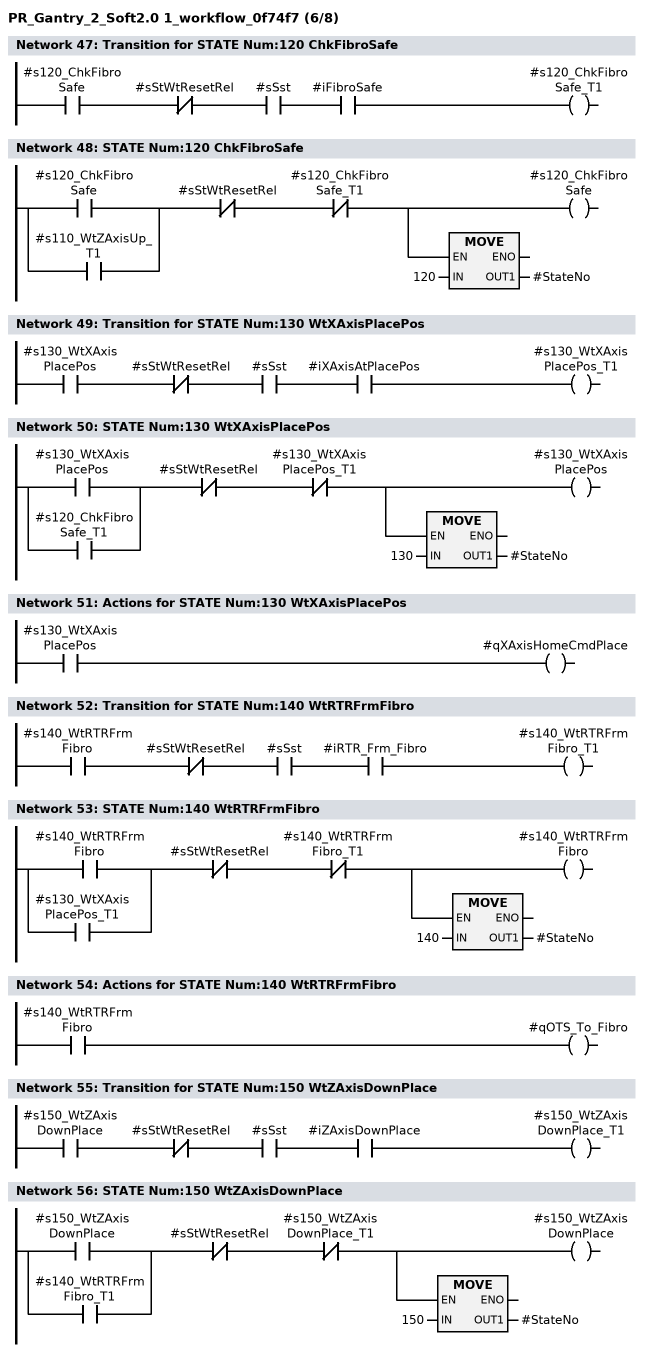
   RUNG wire#powerrail
      Contact( #s120_ChkFibroSafe )
      I_Contact( #sStWtResetRel )
      Contact( #sSst )
      Contact( #iFibroSafe )
      Coil( #s120_ChkFibroSafe_T1 )
   END_RUNG
   // the same network as SCL:
   #s120_ChkFibroSafe_T1 := #s120_ChkFibroSafe AND NOT #sStWtResetRel AND #sSst AND #iFibroSafe;
END_REGION

REGION Network 48: STATE Num:120 ChkFibroSafe
   RUNG wire#powerrail
      Contact( #s120_ChkFibroSafe )
      wire#w1
      I_Contact( #sStWtResetRel )
      I_Contact( #s120_ChkFibroSafe_T1 )
      wire#w2
      Coil( #s120_ChkFibroSafe )
   END_RUNG
   RUNG wire#powerrail
      Contact( #s110_WtZAxisUp_T1 )
   END_RUNG wire#w1
   RUNG wire#w2
      { S7_GenerateENO := "TRUE" } Move(in := 120, out1 => #StateNo)
   END_RUNG
   // the same network as SCL:
   #s120_ChkFibroSafe := (#s120_ChkFibroSafe OR #s110_WtZAxisUp_T1) AND NOT #sStWtResetRel AND NOT #s120_ChkFibroSafe_T1;
   IF #s120_ChkFibroSafe THEN #StateNo := 120; END_IF;
END_REGION

REGION Network 49: Transition for STATE Num:130 WtXAxisPlacePos
   RUNG wire#powerrail
      Contact( #s130_WtXAxisPlacePos )
      I_Contact( #sStWtResetRel )
      Contact( #sSst )
      Contact( #iXAxisAtPlacePos )
      Coil( #s130_WtXAxisPlacePos_T1 )
   END_RUNG
   // the same network as SCL:
   #s130_WtXAxisPlacePos_T1 := #s130_WtXAxisPlacePos AND NOT #sStWtResetRel AND #sSst AND #iXAxisAtPlacePos;
END_REGION

REGION Network 50: STATE Num:130 WtXAxisPlacePos
   RUNG wire#powerrail
      Contact( #s130_WtXAxisPlacePos )
      wire#w1
      I_Contact( #sStWtResetRel )
      I_Contact( #s130_WtXAxisPlacePos_T1 )
      wire#w2
      Coil( #s130_WtXAxisPlacePos )
   END_RUNG
   RUNG wire#powerrail
      Contact( #s120_ChkFibroSafe_T1 )
   END_RUNG wire#w1
   RUNG wire#w2
      { S7_GenerateENO := "TRUE" } Move(in := 130, out1 => #StateNo)
   END_RUNG
   // the same network as SCL:
   #s130_WtXAxisPlacePos := (#s130_WtXAxisPlacePos OR #s120_ChkFibroSafe_T1) AND NOT #sStWtResetRel AND NOT #s130_WtXAxisPlacePos_T1;
   IF #s130_WtXAxisPlacePos THEN #StateNo := 130; END_IF;
END_REGION

REGION Network 51: Actions for STATE Num:130 WtXAxisPlacePos
   RUNG wire#powerrail
      Contact( #s130_WtXAxisPlacePos )
      Coil( #qXAxisHomeCmdPlace )
   END_RUNG
   // the same network as SCL:
   #qXAxisHomeCmdPlace := #s130_WtXAxisPlacePos;
END_REGION

REGION Network 52: Transition for STATE Num:140 WtRTRFrmFibro
   RUNG wire#powerrail
      Contact( #s140_WtRTRFrmFibro )
      I_Contact( #sStWtResetRel )
      Contact( #sSst )
      Contact( #iRTR_Frm_Fibro )
      Coil( #s140_WtRTRFrmFibro_T1 )
   END_RUNG
   // the same network as SCL:
   #s140_WtRTRFrmFibro_T1 := #s140_WtRTRFrmFibro AND NOT #sStWtResetRel AND #sSst AND #iRTR_Frm_Fibro;
END_REGION

REGION Network 53: STATE Num:140 WtRTRFrmFibro
   RUNG wire#powerrail
      Contact( #s140_WtRTRFrmFibro )
      wire#w1
      I_Contact( #sStWtResetRel )
      I_Contact( #s140_WtRTRFrmFibro_T1 )
      wire#w2
      Coil( #s140_WtRTRFrmFibro )
   END_RUNG
   RUNG wire#powerrail
      Contact( #s130_WtXAxisPlacePos_T1 )
   END_RUNG wire#w1
   RUNG wire#w2
      { S7_GenerateENO := "TRUE" } Move(in := 140, out1 => #StateNo)
   END_RUNG
   // the same network as SCL:
   #s140_WtRTRFrmFibro := (#s140_WtRTRFrmFibro OR #s130_WtXAxisPlacePos_T1) AND NOT #sStWtResetRel AND NOT #s140_WtRTRFrmFibro_T1;
   IF #s140_WtRTRFrmFibro THEN #StateNo := 140; END_IF;
END_REGION

REGION Network 54: Actions for STATE Num:140 WtRTRFrmFibro
   RUNG wire#powerrail
      Contact( #s140_WtRTRFrmFibro )
      Coil( #qOTS_To_Fibro )
   END_RUNG
   // the same network as SCL:
   #qOTS_To_Fibro := #s140_WtRTRFrmFibro;
END_REGION

REGION Network 55: Transition for STATE Num:150 WtZAxisDownPlace
   RUNG wire#powerrail
      Contact( #s150_WtZAxisDownPlace )
      I_Contact( #sStWtResetRel )
      Contact( #sSst )
      Contact( #iZAxisDownPlace )
      Coil( #s150_WtZAxisDownPlace_T1 )
   END_RUNG
   // the same network as SCL:
   #s150_WtZAxisDownPlace_T1 := #s150_WtZAxisDownPlace AND NOT #sStWtResetRel AND #sSst AND #iZAxisDownPlace;
END_REGION

REGION Network 56: STATE Num:150 WtZAxisDownPlace
   RUNG wire#powerrail
      Contact( #s150_WtZAxisDownPlace )
      wire#w1
      I_Contact( #sStWtResetRel )
      I_Contact( #s150_WtZAxisDownPlace_T1 )
      wire#w2
      Coil( #s150_WtZAxisDownPlace )
   END_RUNG
   RUNG wire#powerrail
      Contact( #s140_WtRTRFrmFibro_T1 )
   END_RUNG wire#w1
   RUNG wire#w2
      { S7_GenerateENO := "TRUE" } Move(in := 150, out1 => #StateNo)
   END_RUNG
   // the same network as SCL:
   #s150_WtZAxisDownPlace := (#s150_WtZAxisDownPlace OR #s140_WtRTRFrmFibro_T1) AND NOT #sStWtResetRel AND NOT #s150_WtZAxisDownPlace_T1;
   IF #s150_WtZAxisDownPlace THEN #StateNo := 150; END_IF;
END_REGION

REGION Network 57: Actions for STATE Num:150 WtZAxisDownPlace
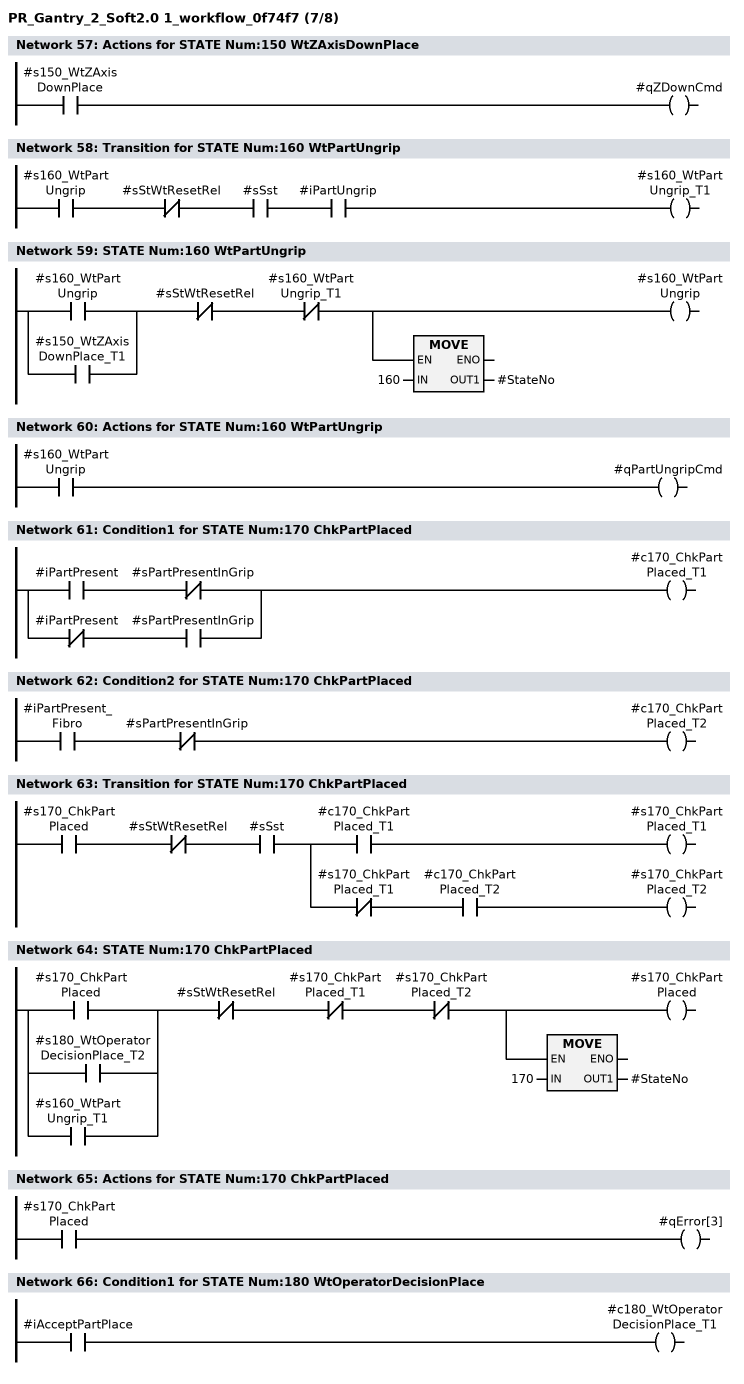
   RUNG wire#powerrail
      Contact( #s150_WtZAxisDownPlace )
      Coil( #qZDownCmd )
   END_RUNG
   // the same network as SCL:
   #qZDownCmd := #s150_WtZAxisDownPlace;
END_REGION

REGION Network 58: Transition for STATE Num:160 WtPartUngrip
   RUNG wire#powerrail
      Contact( #s160_WtPartUngrip )
      I_Contact( #sStWtResetRel )
      Contact( #sSst )
      Contact( #iPartUngrip )
      Coil( #s160_WtPartUngrip_T1 )
   END_RUNG
   // the same network as SCL:
   #s160_WtPartUngrip_T1 := #s160_WtPartUngrip AND NOT #sStWtResetRel AND #sSst AND #iPartUngrip;
END_REGION

REGION Network 59: STATE Num:160 WtPartUngrip
   RUNG wire#powerrail
      Contact( #s160_WtPartUngrip )
      wire#w1
      I_Contact( #sStWtResetRel )
      I_Contact( #s160_WtPartUngrip_T1 )
      wire#w2
      Coil( #s160_WtPartUngrip )
   END_RUNG
   RUNG wire#powerrail
      Contact( #s150_WtZAxisDownPlace_T1 )
   END_RUNG wire#w1
   RUNG wire#w2
      { S7_GenerateENO := "TRUE" } Move(in := 160, out1 => #StateNo)
   END_RUNG
   // the same network as SCL:
   #s160_WtPartUngrip := (#s160_WtPartUngrip OR #s150_WtZAxisDownPlace_T1) AND NOT #sStWtResetRel AND NOT #s160_WtPartUngrip_T1;
   IF #s160_WtPartUngrip THEN #StateNo := 160; END_IF;
END_REGION

REGION Network 60: Actions for STATE Num:160 WtPartUngrip
   RUNG wire#powerrail
      Contact( #s160_WtPartUngrip )
      Coil( #qPartUngripCmd )
   END_RUNG
   // the same network as SCL:
   #qPartUngripCmd := #s160_WtPartUngrip;
END_REGION

REGION Network 61: Condition1 for STATE Num:170 ChkPartPlaced
   RUNG wire#powerrail
      Contact( #iPartPresent )
      I_Contact( #sPartPresentInGrip )
      wire#w1
      Coil( #c170_ChkPartPlaced_T1 )
   END_RUNG
   RUNG wire#powerrail
      I_Contact( #iPartPresent )
      Contact( #sPartPresentInGrip )
   END_RUNG wire#w1
   // the same network as SCL:
   #c170_ChkPartPlaced_T1 := (#iPartPresent AND NOT #sPartPresentInGrip) OR (NOT #iPartPresent AND #sPartPresentInGrip);
END_REGION

REGION Network 62: Condition2 for STATE Num:170 ChkPartPlaced
   RUNG wire#powerrail
      Contact( #iPartPresent_Fibro )
      I_Contact( #sPartPresentInGrip )
      Coil( #c170_ChkPartPlaced_T2 )
   END_RUNG
   // the same network as SCL:
   #c170_ChkPartPlaced_T2 := #iPartPresent_Fibro AND NOT #sPartPresentInGrip;
END_REGION

REGION Network 63: Transition for STATE Num:170 ChkPartPlaced
   RUNG wire#powerrail
      Contact( #s170_ChkPartPlaced )
      I_Contact( #sStWtResetRel )
      Contact( #sSst )
      wire#w1
      Contact( #c170_ChkPartPlaced_T1 )
      Coil( #s170_ChkPartPlaced_T1 )
   END_RUNG
   RUNG wire#w1
      I_Contact( #s170_ChkPartPlaced_T1 )
      Contact( #c170_ChkPartPlaced_T2 )
      Coil( #s170_ChkPartPlaced_T2 )
   END_RUNG
   // the same network as SCL:
   #_w1 := #s170_ChkPartPlaced AND NOT #sStWtResetRel AND #sSst;
   #s170_ChkPartPlaced_T1 := #_w1 AND #c170_ChkPartPlaced_T1;
   #s170_ChkPartPlaced_T2 := #_w1 AND NOT #s170_ChkPartPlaced_T1 AND #c170_ChkPartPlaced_T2;
END_REGION

REGION Network 64: STATE Num:170 ChkPartPlaced
   RUNG wire#powerrail
      Contact( #s170_ChkPartPlaced )
      wire#w1
      I_Contact( #sStWtResetRel )
      I_Contact( #s170_ChkPartPlaced_T1 )
      I_Contact( #s170_ChkPartPlaced_T2 )
      wire#w2
      Coil( #s170_ChkPartPlaced )
   END_RUNG
   RUNG wire#powerrail
      Contact( #s180_WtOperatorDecisionPlace_T2 )
   END_RUNG wire#w1
   RUNG wire#powerrail
      Contact( #s160_WtPartUngrip_T1 )
   END_RUNG wire#w1
   RUNG wire#w2
      { S7_GenerateENO := "TRUE" } Move(in := 170, out1 => #StateNo)
   END_RUNG
   // the same network as SCL:
   #s170_ChkPartPlaced := (#s170_ChkPartPlaced OR #s180_WtOperatorDecisionPlace_T2 OR #s160_WtPartUngrip_T1) AND NOT #sStWtResetRel AND NOT #s170_ChkPartPlaced_T1 AND NOT #s170_ChkPartPlaced_T2;
   IF #s170_ChkPartPlaced THEN #StateNo := 170; END_IF;
END_REGION

REGION Network 65: Actions for STATE Num:170 ChkPartPlaced
   RUNG wire#powerrail
      Contact( #s170_ChkPartPlaced )
      Coil( #qError[3] )
   END_RUNG
   // the same network as SCL:
   #qError[3] := #s170_ChkPartPlaced;
END_REGION

REGION Network 66: Condition1 for STATE Num:180 WtOperatorDecisionPlace
   RUNG wire#powerrail
      Contact( #iAcceptPartPlace )
      Coil( #c180_WtOperatorDecisionPlace_T1 )
   END_RUNG
   // the same network as SCL:
   #c180_WtOperatorDecisionPlace_T1 := #iAcceptPartPlace;
END_REGION

REGION Network 67: Condition2 for STATE Num:180 WtOperatorDecisionPlace
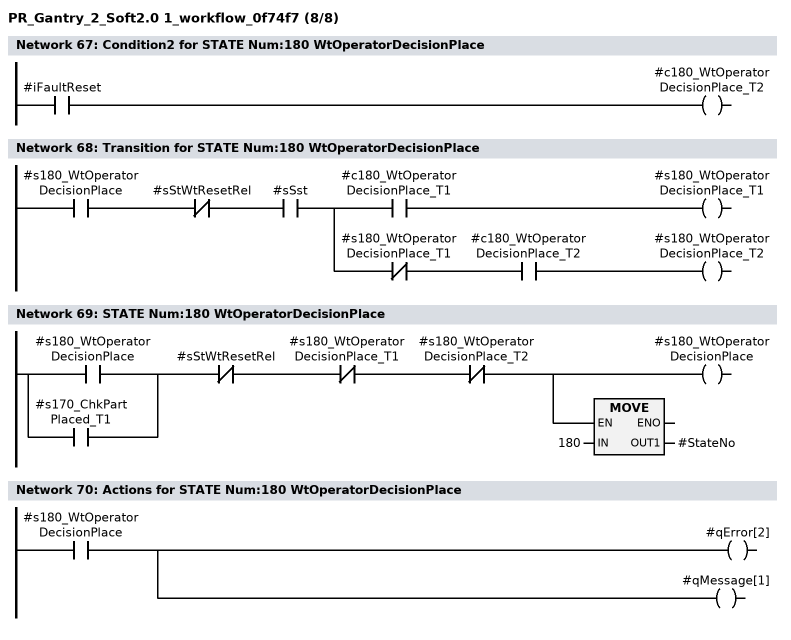
   RUNG wire#powerrail
      Contact( #iFaultReset )
      Coil( #c180_WtOperatorDecisionPlace_T2 )
   END_RUNG
   // the same network as SCL:
   #c180_WtOperatorDecisionPlace_T2 := #iFaultReset;
END_REGION

REGION Network 68: Transition for STATE Num:180 WtOperatorDecisionPlace
   RUNG wire#powerrail
      Contact( #s180_WtOperatorDecisionPlace )
      I_Contact( #sStWtResetRel )
      Contact( #sSst )
      wire#w1
      Contact( #c180_WtOperatorDecisionPlace_T1 )
      Coil( #s180_WtOperatorDecisionPlace_T1 )
   END_RUNG
   RUNG wire#w1
      I_Contact( #s180_WtOperatorDecisionPlace_T1 )
      Contact( #c180_WtOperatorDecisionPlace_T2 )
      Coil( #s180_WtOperatorDecisionPlace_T2 )
   END_RUNG
   // the same network as SCL:
   #_w1 := #s180_WtOperatorDecisionPlace AND NOT #sStWtResetRel AND #sSst;
   #s180_WtOperatorDecisionPlace_T1 := #_w1 AND #c180_WtOperatorDecisionPlace_T1;
   #s180_WtOperatorDecisionPlace_T2 := #_w1 AND NOT #s180_WtOperatorDecisionPlace_T1 AND #c180_WtOperatorDecisionPlace_T2;
END_REGION

REGION Network 69: STATE Num:180 WtOperatorDecisionPlace
   RUNG wire#powerrail
      Contact( #s180_WtOperatorDecisionPlace )
      wire#w1
      I_Contact( #sStWtResetRel )
      I_Contact( #s180_WtOperatorDecisionPlace_T1 )
      I_Contact( #s180_WtOperatorDecisionPlace_T2 )
      wire#w2
      Coil( #s180_WtOperatorDecisionPlace )
   END_RUNG
   RUNG wire#powerrail
      Contact( #s170_ChkPartPlaced_T1 )
   END_RUNG wire#w1
   RUNG wire#w2
      { S7_GenerateENO := "TRUE" } Move(in := 180, out1 => #StateNo)
   END_RUNG
   // the same network as SCL:
   #s180_WtOperatorDecisionPlace := (#s180_WtOperatorDecisionPlace OR #s170_ChkPartPlaced_T1) AND NOT #sStWtResetRel AND NOT #s180_WtOperatorDecisionPlace_T1 AND NOT #s180_WtOperatorDecisionPlace_T2;
   IF #s180_WtOperatorDecisionPlace THEN #StateNo := 180; END_IF;
END_REGION

REGION Network 70: Actions for STATE Num:180 WtOperatorDecisionPlace
   RUNG wire#powerrail
      Contact( #s180_WtOperatorDecisionPlace )
      wire#w1
      Coil( #qError[2] )
   END_RUNG
   RUNG wire#w1
      Coil( #qMessage[1] )
   END_RUNG
   // the same network as SCL:
   #qError[2] := #s180_WtOperatorDecisionPlace;
   #qMessage[1] := #s180_WtOperatorDecisionPlace;
END_REGION
END_FUNCTION_BLOCK
